(* IEC 61131-3 sources: Repository_IEMA_Test/LMC_PacDrive.device.xml.v3^/Plc Logic.plclogic.xml.v3^/Application.application.xml.v3^/TemplateFullProgrammingFramework/Examples/ExampleModulesExtItf/FB_AxisModuleExtItf.fb.st^, 1 file *)

(* ---- RegisterLoggerPoint.meth.st ---- *)
METHOD PUBLIC RegisterLoggerPoint
VAR_INPUT
	i_ifParent		: APL.IF_LoggerPoint;
	i_sName			: STRING[80];
END_VAR
VAR_OUTPUT
	q_etDiag		: GD.ET_Diag := GD.ET_Diag.Ok;
	q_etDiagExt		: AXM.ET_DiagExt := AXM.ET_DiagExt.Ok;
END_VAR

THIS^.fbAxisModule.RegisterLoggerPoint(	i_ifParent	:= i_ifParent,
										i_sName		:= i_sName,
										q_etDiag	=> q_etDiag,
										q_etDiagExt	=> q_etDiagExt);
